// Mitsubishi GX Works2 project: FINAL_V7   PLC: Q03UDV

PROGRAM MAIN
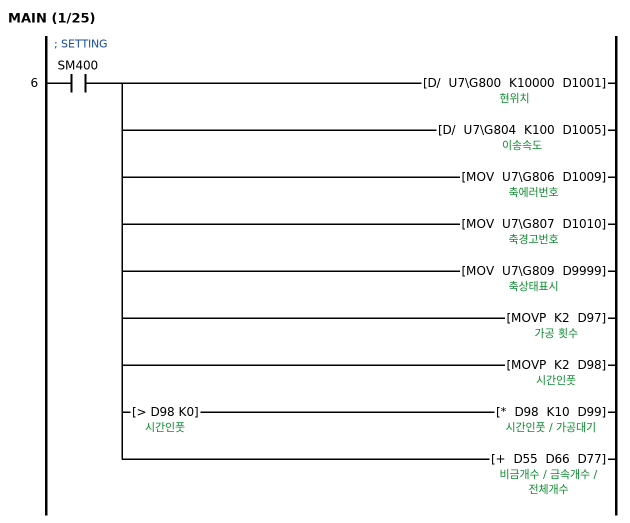
; SETTING
6     LD      SM400
      D/      U7\G800 K10000 D1001  ; 현위치
      D/      U7\G804 K100 D1005  ; 이송속도
      MOV     U7\G806 D1009  ; 축에러번호
      MOV     U7\G807 D1010  ; 축경고번호
      MOV     U7\G809 D9999  ; 축상태표시
      MOVP    K2 D97  ; 가공 횟수
      MOVP    K2 D98  ; 시간인풋
      MPS
      AND>    D98 K0  ; 시간인풋
      *       D98 K10 D99  ; 가공대기
      MPP
      +       D55 D66 D77  ; 비금개수 / 금속개수 / 전체개수
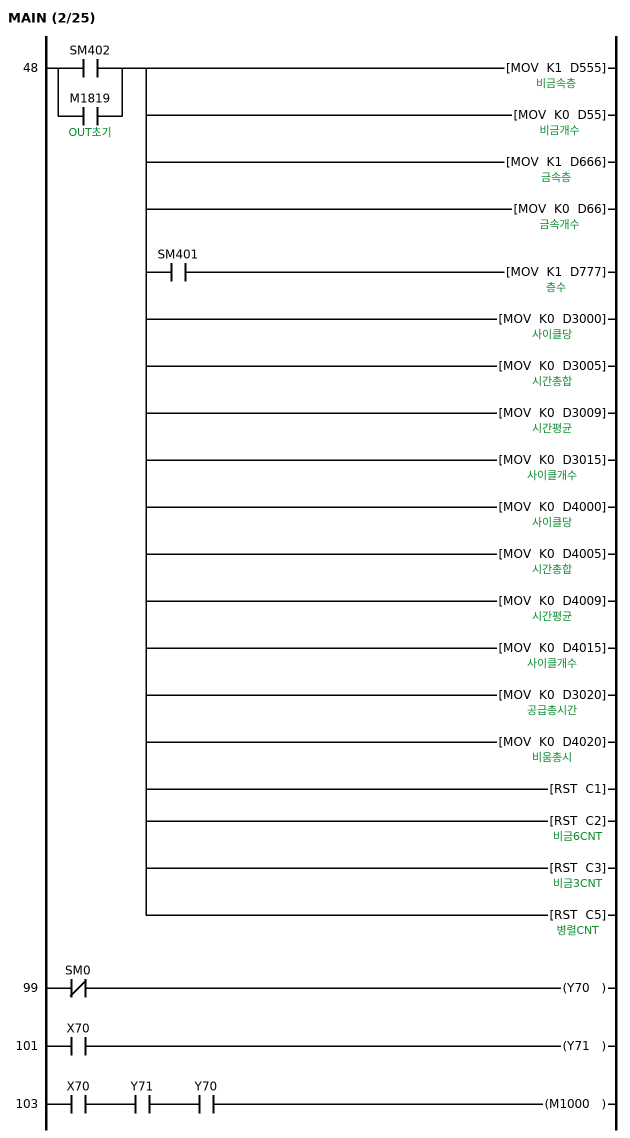
48    LD      SM402
      OR      M1819  ; OUT초기
      MOV     K1 D555  ; 비금속층
      MOV     K0 D55
      MOV     K1 D666  ; 금속층
      MOV     K0 D66
      MPS
      AND     SM401
      MOV     K1 D777  ; 층수
      MPP
      MOV     K0 D3000  ; 사이클당
      MOV     K0 D3005  ; 시간총합
      MOV     K0 D3009  ; 시간평균
      MOV     K0 D3015  ; 사이클개수
      MOV     K0 D4000  ; 사이클당
      MOV     K0 D4005  ; 시간총합
      MOV     K0 D4009  ; 시간평균
      MOV     K0 D4015  ; 사이클개수
      MOV     K0 D3020  ; 공급총시간
      MOV     K0 D4020  ; 비움총시
      RST     C1
      RST     C2  ; 비금6CNT
      RST     C3  ; 비금3CNT
      RST     C5  ; 병렬CNT
99    LDI     SM0
      OUT     Y70
101   LD      X70
      OUT     Y71
103   LD      X70
      AND     Y71
      AND     Y70
      OUT     M1000
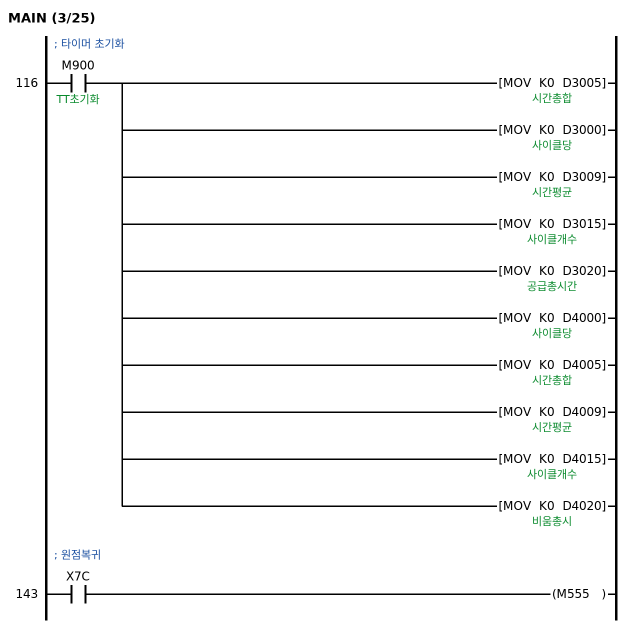
; 타이머 초기화
116   LD      M900  ; TT초기화
      MOV     K0 D3005
      MOV     K0 D3000
      MOV     K0 D3009
      MOV     K0 D3015
      MOV     K0 D3020
      MOV     K0 D4000
      MOV     K0 D4005
      MOV     K0 D4009
      MOV     K0 D4015
      MOV     K0 D4020
; 원점복귀
143   LD      X7C
      OUT     M555
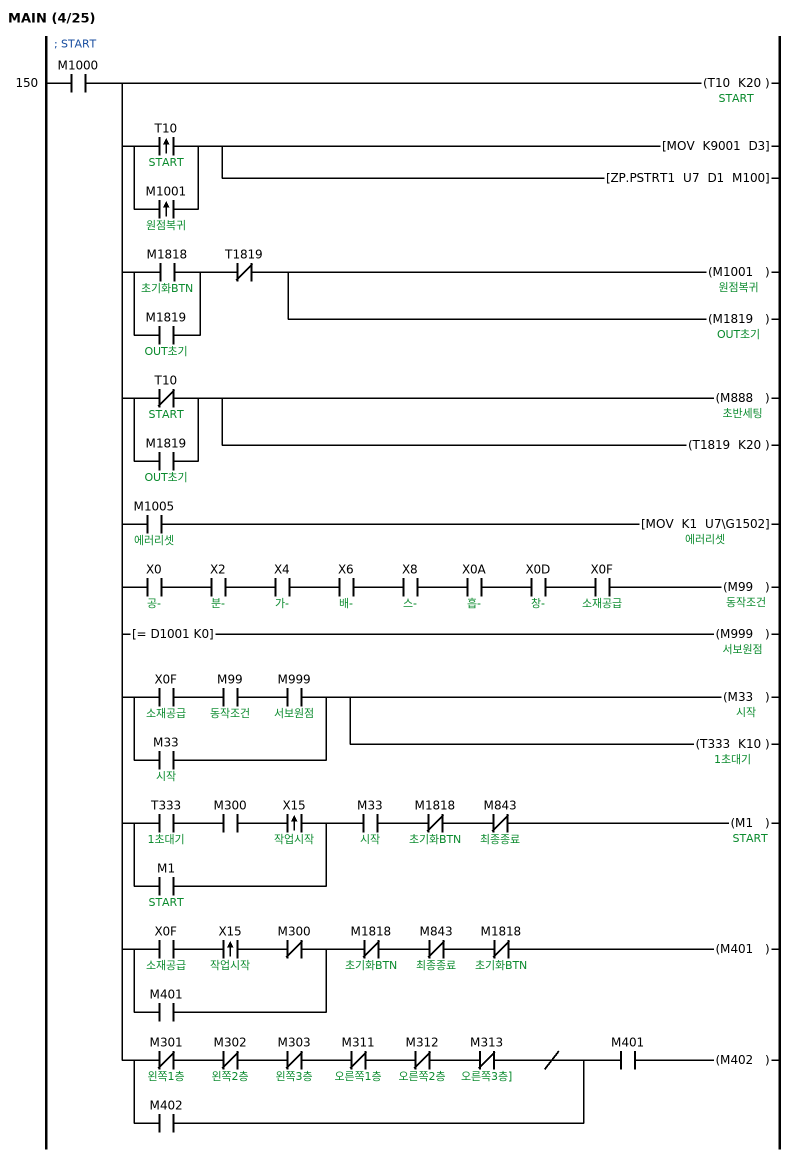
; START
150   LD      M1000
      OUT     T10 K20  ; START
      MPS
      LDP     T10  ; START
      ORP     M1001  ; 원점복귀
      ANB
      MOV     K9001 D3
      ZP.PSTRT1 U7 D1 M100
      MRD
      LD      M1818  ; 초기화BTN
      OR      M1819  ; OUT초기
      ANB
      ANI     T1819
      OUT     M1001  ; 원점복귀
      OUT     M1819  ; OUT초기
      MRD
      LDI     T10  ; START
      OR      M1819  ; OUT초기
      ANB
      OUT     M888  ; 초반세팅
      OUT     T1819 K20
      MRD
      AND     M1005  ; 에러리셋
      MOV     K1 U7\G1502  ; 에러리셋
      MRD
      AND     X0  ; 공-
      AND     X2  ; 분-
      AND     X4  ; 가-
      AND     X6  ; 배-
      AND     X8  ; 스-
      AND     X0A  ; 흡-
      AND     X0D  ; 창-
      AND     X0F  ; 소재공급
      OUT     M99  ; 동작조건
      MRD
      AND=    D1001 K0
      OUT     M999  ; 서보원점
      MRD
      LD      X0F  ; 소재공급
      AND     M99  ; 동작조건
      AND     M999  ; 서보원점
      OR      M33  ; 시작
      ANB
      OUT     M33  ; 시작
      OUT     T333 K10  ; 1초대기
      MRD
      LD      T333  ; 1초대기
      AND     M300
      ANDP    X15  ; 작업시작
      OR      M1  ; START
      ANB
      AND     M33  ; 시작
      ANI     M1818  ; 초기화BTN
      ANI     M843  ; 최종종료
      OUT     M1  ; START
      MRD
      LD      X0F  ; 소재공급
      ANDP    X15  ; 작업시작
      ANI     M300
      OR      M401
      ANB
      ANI     M1818  ; 초기화BTN
      ANI     M843  ; 최종종료
      ANI     M1818  ; 초기화BTN
      OUT     M401
      MPP
      LDI     M301  ; 왼쪽1층
      ANI     M302  ; 왼쪽2층
      ANI     M303  ; 왼쪽3층
      ANI     M311  ; 오른쪽1층
      ANI     M312  ; 오른쪽2층
      ANI     M313  ; 오른쪽3층]
      INV
      OR      M402
      ANB
      AND     M401
      OUT     M402
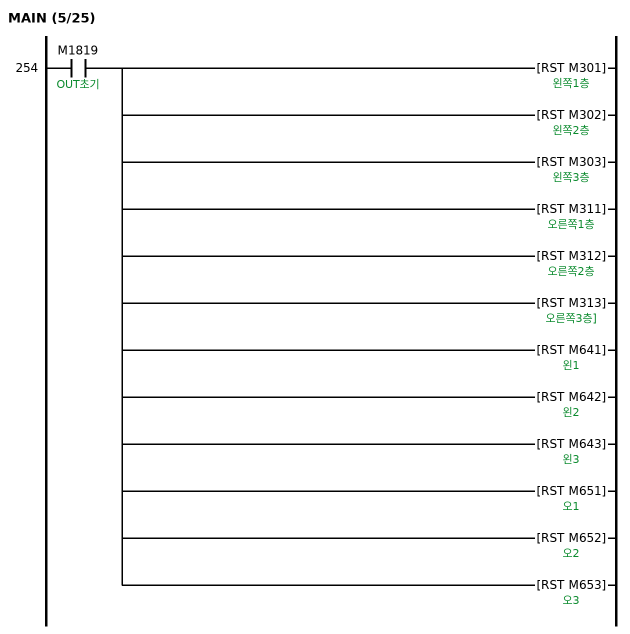
254   LD      M1819  ; OUT초기
      RST     M301  ; 왼쪽1층
      RST     M302  ; 왼쪽2층
      RST     M303  ; 왼쪽3층
      RST     M311  ; 오른쪽1층
      RST     M312  ; 오른쪽2층
      RST     M313  ; 오른쪽3층]
      RST     M641  ; 왼1
      RST     M642  ; 왼2
      RST     M643  ; 왼3
      RST     M651  ; 오1
      RST     M652  ; 오2
      RST     M653  ; 오3
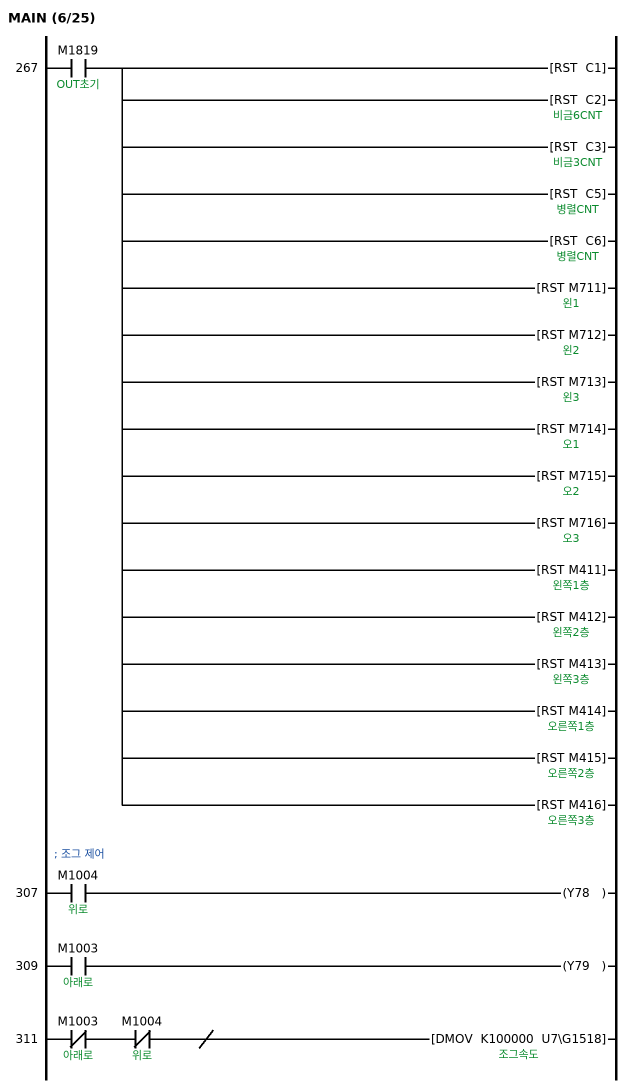
267   LD      M1819  ; OUT초기
      RST     C1
      RST     C2  ; 비금6CNT
      RST     C3  ; 비금3CNT
      RST     C5  ; 병렬CNT
      RST     C6  ; 병렬CNT
      RST     M711  ; 왼1
      RST     M712  ; 왼2
      RST     M713  ; 왼3
      RST     M714  ; 오1
      RST     M715  ; 오2
      RST     M716  ; 오3
      RST     M411  ; 왼쪽1층
      RST     M412  ; 왼쪽2층
      RST     M413  ; 왼쪽3층
      RST     M414  ; 오른쪽1층
      RST     M415  ; 오른쪽2층
      RST     M416  ; 오른쪽3층
; 조그 제어
307   LD      M1004  ; 위로
      OUT     Y78
309   LD      M1003  ; 아래로
      OUT     Y79
311   LDI     M1003  ; 아래로
      ANI     M1004  ; 위로
      INV
      DMOV    K100000 U7\G1518  ; 조그속도
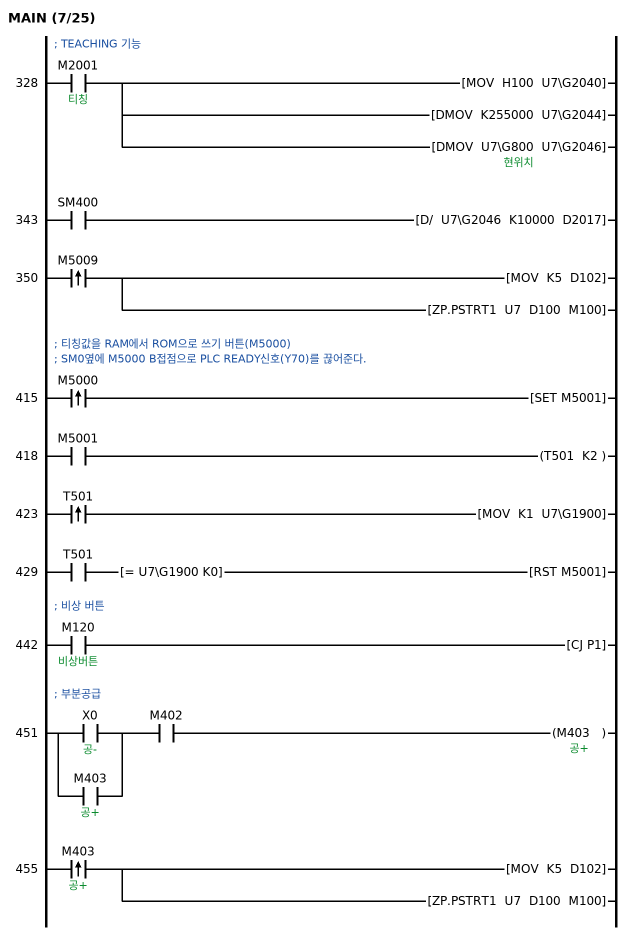
; TEACHING 기능
328   LD      M2001  ; 티칭
      MOV     H100 U7\G2040
      DMOV    K255000 U7\G2044
      DMOV    U7\G800 U7\G2046
343   LD      SM400
      D/      U7\G2046 K10000 D2017
350   LDP     M5009
      MOV     K5 D102
      ZP.PSTRT1 U7 D100 M100
; 티칭값을 RAM에서 ROM으로 쓰기 버튼(M5000)
; SM0옆에 M5000 B접점으로 PLC READY신호(Y70)를 끊어준다.
415   LDP     M5000
      SET     M5001
418   LD      M5001
      OUT     T501 K2
423   LDP     T501
      MOV     K1 U7\G1900
429   LD      T501
      AND=    U7\G1900 K0
      RST     M5001
; 비상 버튼
442   LD      M120  ; 비상버튼
      CJ      P1
; 부분공급
451   LD      X0  ; 공-
      OR      M403  ; 공+
      AND     M402
      OUT     M403  ; 공+
455   LDP     M403  ; 공+
      MOV     K5 D102
      ZP.PSTRT1 U7 D100 M100
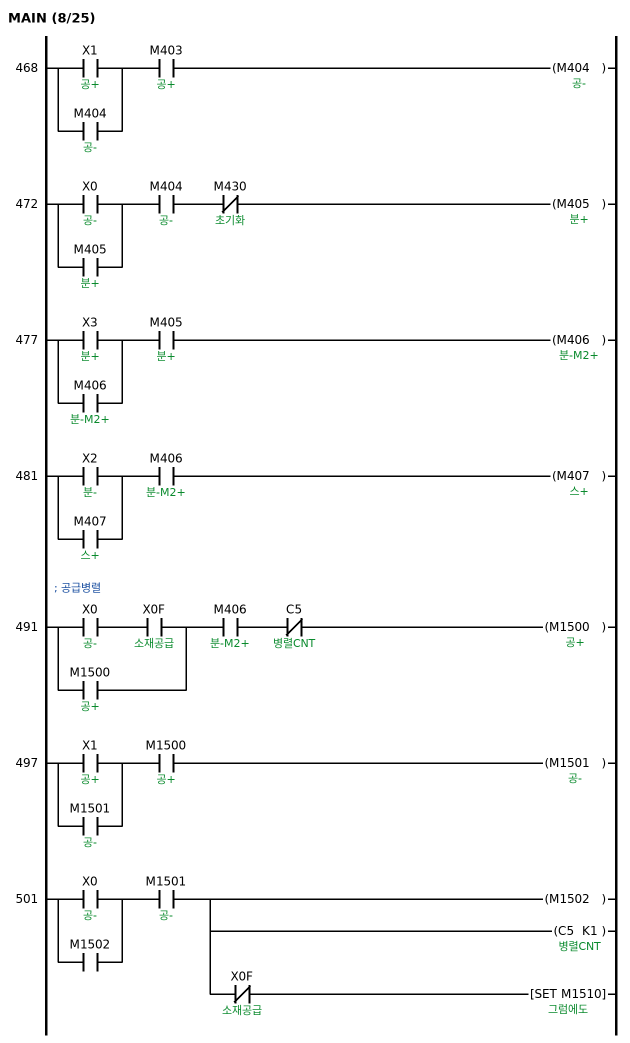
468   LD      X1  ; 공+
      OR      M404  ; 공-
      AND     M403  ; 공+
      OUT     M404  ; 공-
472   LD      X0  ; 공-
      OR      M405  ; 분+
      AND     M404  ; 공-
      ANI     M430  ; 초기화
      OUT     M405  ; 분+
477   LD      X3  ; 분+
      OR      M406  ; 분-M2+
      AND     M405  ; 분+
      OUT     M406  ; 분-M2+
481   LD      X2  ; 분-
      OR      M407  ; 스+
      AND     M406  ; 분-M2+
      OUT     M407  ; 스+
; 공급병렬
491   LD      X0  ; 공-
      AND     X0F  ; 소재공급
      OR      M1500  ; 공+
      AND     M406  ; 분-M2+
      ANI     C5  ; 병렬CNT
      OUT     M1500  ; 공+
497   LD      X1  ; 공+
      OR      M1501  ; 공-
      AND     M1500  ; 공+
      OUT     M1501  ; 공-
501   LD      X0  ; 공-
      OR      M1502
      AND     M1501  ; 공-
      OUT     M1502
      OUT     C5 K1  ; 병렬CNT
      ANI     X0F  ; 소재공급
      SET     M1510  ; 그럼에도
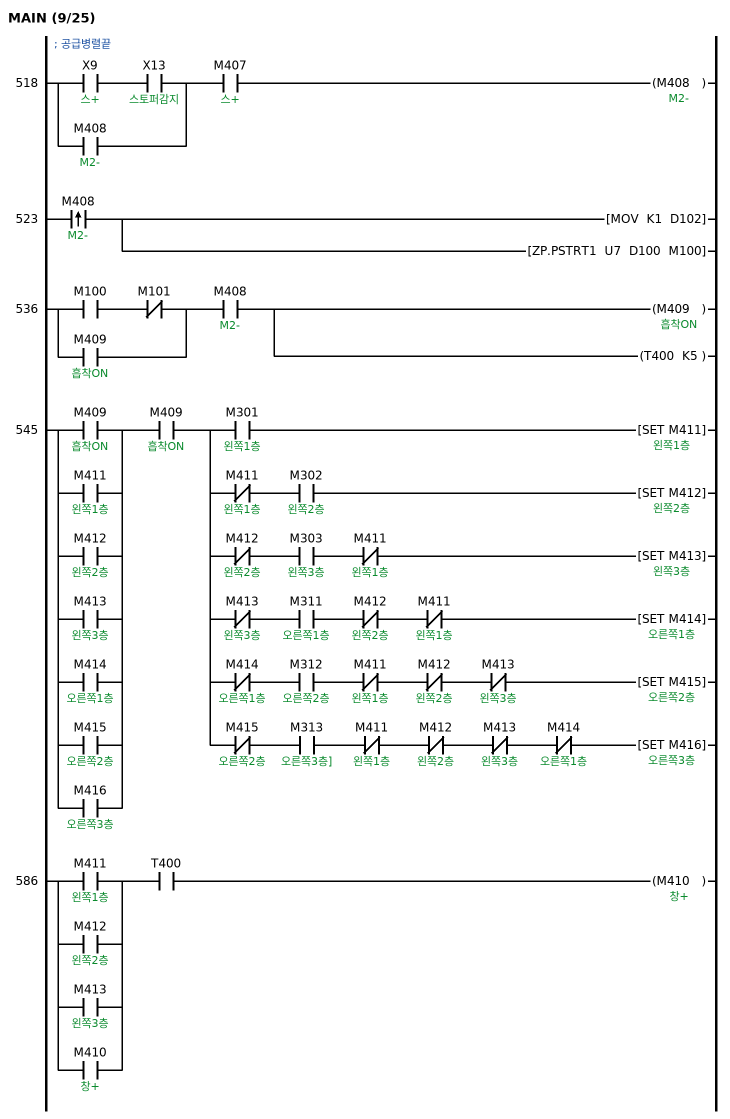
; 공급병렬끝
518   LD      X9  ; 스+
      AND     X13  ; 스토퍼감지
      OR      M408  ; M2-
      AND     M407  ; 스+
      OUT     M408  ; M2-
523   LDP     M408  ; M2-
      MOV     K1 D102
      ZP.PSTRT1 U7 D100 M100
536   LD      M100
      ANI     M101
      OR      M409  ; 흡착ON
      AND     M408  ; M2-
      OUT     M409  ; 흡착ON
      OUT     T400 K5
545   LD      M409  ; 흡착ON
      OR      M411  ; 왼쪽1층
      OR      M412  ; 왼쪽2층
      OR      M413  ; 왼쪽3층
      OR      M414  ; 오른쪽1층
      OR      M415  ; 오른쪽2층
      OR      M416  ; 오른쪽3층
      AND     M409  ; 흡착ON
      MPS
      AND     M301  ; 왼쪽1층
      SET     M411  ; 왼쪽1층
      MRD
      ANI     M411  ; 왼쪽1층
      AND     M302  ; 왼쪽2층
      SET     M412  ; 왼쪽2층
      MRD
      ANI     M412  ; 왼쪽2층
      AND     M303  ; 왼쪽3층
      ANI     M411  ; 왼쪽1층
      SET     M413  ; 왼쪽3층
      MRD
      ANI     M413  ; 왼쪽3층
      AND     M311  ; 오른쪽1층
      ANI     M412  ; 왼쪽2층
      ANI     M411  ; 왼쪽1층
      SET     M414  ; 오른쪽1층
      MRD
      ANI     M414  ; 오른쪽1층
      AND     M312  ; 오른쪽2층
      ANI     M411  ; 왼쪽1층
      ANI     M412  ; 왼쪽2층
      ANI     M413  ; 왼쪽3층
      SET     M415  ; 오른쪽2층
      MPP
      ANI     M415  ; 오른쪽2층
      AND     M313  ; 오른쪽3층]
      ANI     M411  ; 왼쪽1층
      ANI     M412  ; 왼쪽2층
      ANI     M413  ; 왼쪽3층
      ANI     M414  ; 오른쪽1층
      SET     M416  ; 오른쪽3층
586   LD      M411  ; 왼쪽1층
      OR      M412  ; 왼쪽2층
      OR      M413  ; 왼쪽3층
      OR      M410  ; 창+
      AND     T400
      OUT     M410  ; 창+
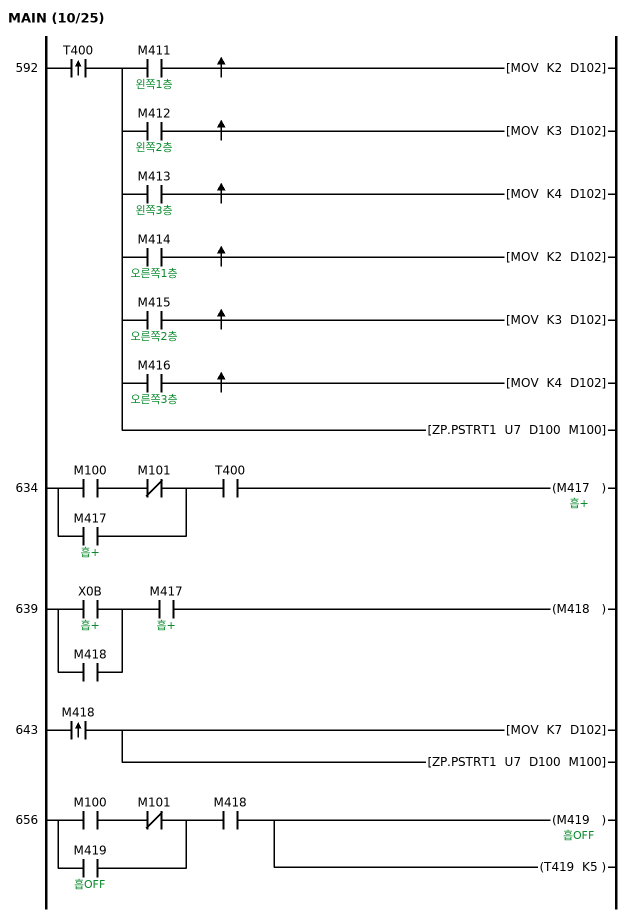
592   LDP     T400
      MPS
      AND     M411  ; 왼쪽1층
      MEP
      MOV     K2 D102
      MRD
      AND     M412  ; 왼쪽2층
      MEP
      MOV     K3 D102
      MRD
      AND     M413  ; 왼쪽3층
      MEP
      MOV     K4 D102
      MRD
      AND     M414  ; 오른쪽1층
      MEP
      MOV     K2 D102
      MRD
      AND     M415  ; 오른쪽2층
      MEP
      MOV     K3 D102
      MRD
      AND     M416  ; 오른쪽3층
      MEP
      MOV     K4 D102
      MPP
      ZP.PSTRT1 U7 D100 M100
634   LD      M100
      ANI     M101
      OR      M417  ; 흡+
      AND     T400
      OUT     M417  ; 흡+
639   LD      X0B  ; 흡+
      OR      M418
      AND     M417  ; 흡+
      OUT     M418
643   LDP     M418
      MOV     K7 D102
      ZP.PSTRT1 U7 D100 M100
656   LD      M100
      ANI     M101
      OR      M419  ; 흡OFF
      AND     M418
      OUT     M419  ; 흡OFF
      OUT     T419 K5
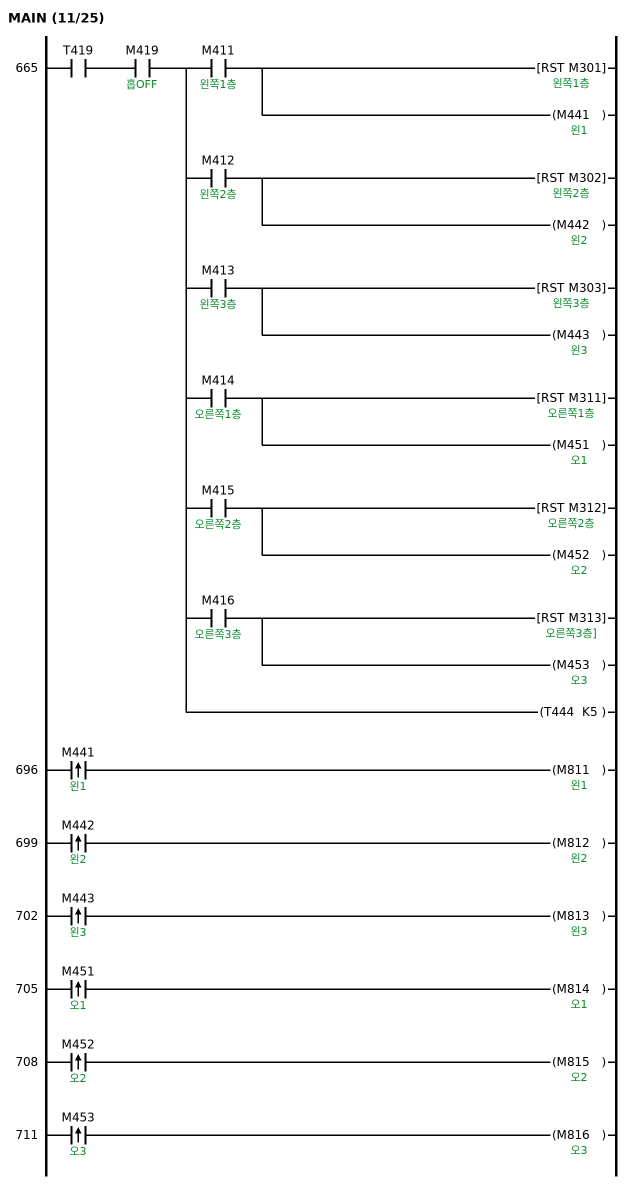
665   LD      T419
      AND     M419  ; 흡OFF
      MPS
      AND     M411  ; 왼쪽1층
      RST     M301  ; 왼쪽1층
      OUT     M441  ; 왼1
      MRD
      AND     M412  ; 왼쪽2층
      RST     M302  ; 왼쪽2층
      OUT     M442  ; 왼2
      MRD
      AND     M413  ; 왼쪽3층
      RST     M303  ; 왼쪽3층
      OUT     M443  ; 왼3
      MRD
      AND     M414  ; 오른쪽1층
      RST     M311  ; 오른쪽1층
      OUT     M451  ; 오1
      MRD
      AND     M415  ; 오른쪽2층
      RST     M312  ; 오른쪽2층
      OUT     M452  ; 오2
      MRD
      AND     M416  ; 오른쪽3층
      RST     M313  ; 오른쪽3층]
      OUT     M453  ; 오3
      MPP
      OUT     T444 K5
696   LDP     M441  ; 왼1
      OUT     M811  ; 왼1
699   LDP     M442  ; 왼2
      OUT     M812  ; 왼2
702   LDP     M443  ; 왼3
      OUT     M813  ; 왼3
705   LDP     M451  ; 오1
      OUT     M814  ; 오1
708   LDP     M452  ; 오2
      OUT     M815  ; 오2
711   LDP     M453  ; 오3
      OUT     M816  ; 오3
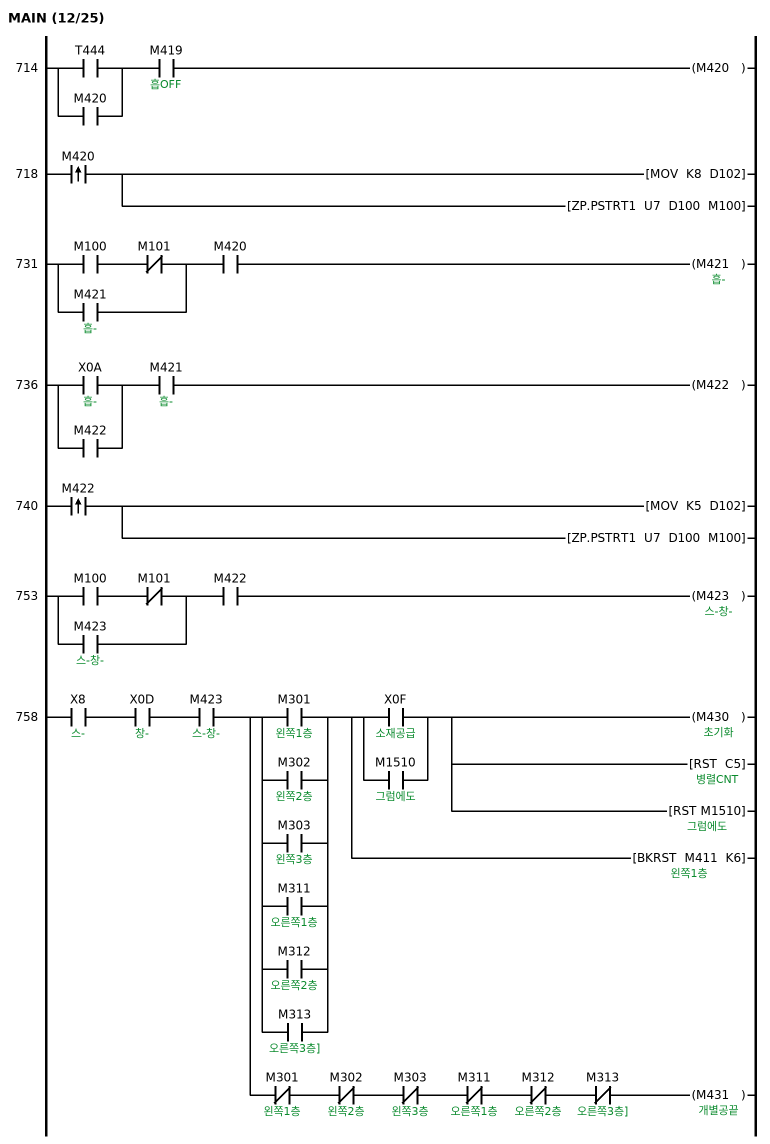
714   LD      T444
      OR      M420
      AND     M419  ; 흡OFF
      OUT     M420
718   LDP     M420
      MOV     K8 D102
      ZP.PSTRT1 U7 D100 M100
731   LD      M100
      ANI     M101
      OR      M421  ; 흡-
      AND     M420
      OUT     M421  ; 흡-
736   LD      X0A  ; 흡-
      OR      M422
      AND     M421  ; 흡-
      OUT     M422
740   LDP     M422
      MOV     K5 D102
      ZP.PSTRT1 U7 D100 M100
753   LD      M100
      ANI     M101
      OR      M423  ; 스-창-
      AND     M422
      OUT     M423  ; 스-창-
758   LD      X8  ; 스-
      AND     X0D  ; 창-
      AND     M423  ; 스-창-
      MPS
      LD      M301  ; 왼쪽1층
      OR      M302  ; 왼쪽2층
      OR      M303  ; 왼쪽3층
      OR      M311  ; 오른쪽1층
      OR      M312  ; 오른쪽2층
      OR      M313  ; 오른쪽3층]
      ANB
      MPS
      LD      X0F  ; 소재공급
      OR      M1510  ; 그럼에도
      ANB
      OUT     M430  ; 초기화
      RST     C5  ; 병렬CNT
      RST     M1510  ; 그럼에도
      MPP
      BKRST   M411 K6
      MPP
      ANI     M301  ; 왼쪽1층
      ANI     M302  ; 왼쪽2층
      ANI     M303  ; 왼쪽3층
      ANI     M311  ; 오른쪽1층
      ANI     M312  ; 오른쪽2층
      ANI     M313  ; 오른쪽3층]
      OUT     M431  ; 개별공끝
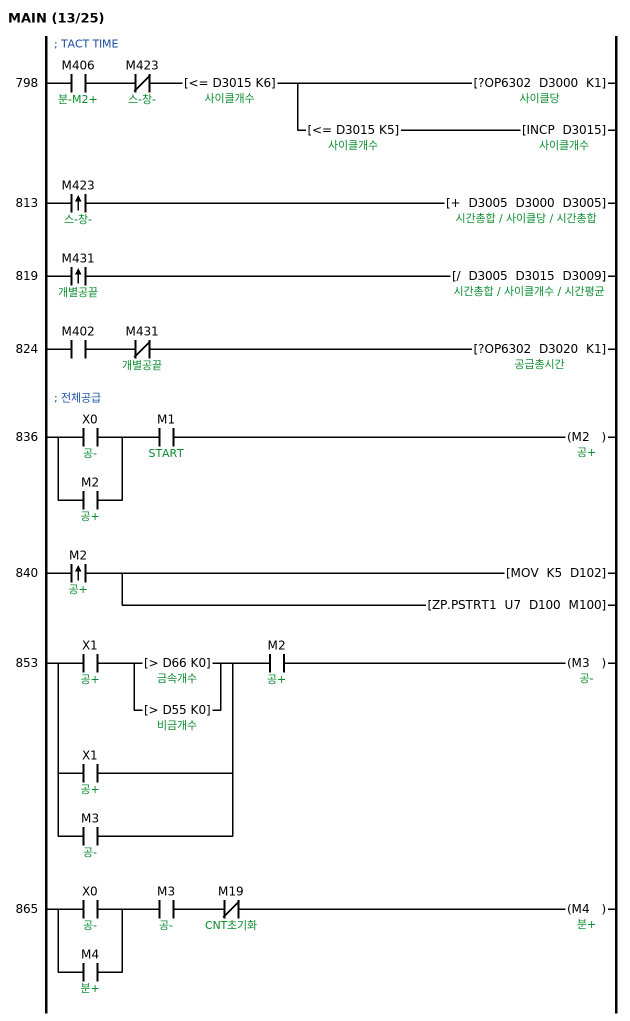
; TACT TIME
798   LD      M406  ; 분-M2+
      ANI     M423  ; 스-창-
      AND<=   D3015 K6  ; 사이클개수
      ?OP6302 D3000 K1
      AND<=   D3015 K5  ; 사이클개수
      INCP    D3015
813   LDP     M423  ; 스-창-
      +       D3005 D3000 D3005
819   LDP     M431  ; 개별공끝
      /       D3005 D3015 D3009
824   LD      M402
      ANI     M431  ; 개별공끝
      ?OP6302 D3020 K1
; 전체공급
836   LD      X0  ; 공-
      OR      M2  ; 공+
      AND     M1  ; START
      OUT     M2  ; 공+
840   LDP     M2  ; 공+
      MOV     K5 D102
      ZP.PSTRT1 U7 D100 M100
853   LD      X1  ; 공+
      LD>     D66 K0  ; 금속개수
      OR>     D55 K0  ; 비금개수
      ANB
      OR      X1  ; 공+
      OR      M3  ; 공-
      AND     M2  ; 공+
      OUT     M3  ; 공-
865   LD      X0  ; 공-
      OR      M4  ; 분+
      AND     M3  ; 공-
      ANI     M19  ; CNT초기화
      OUT     M4  ; 분+
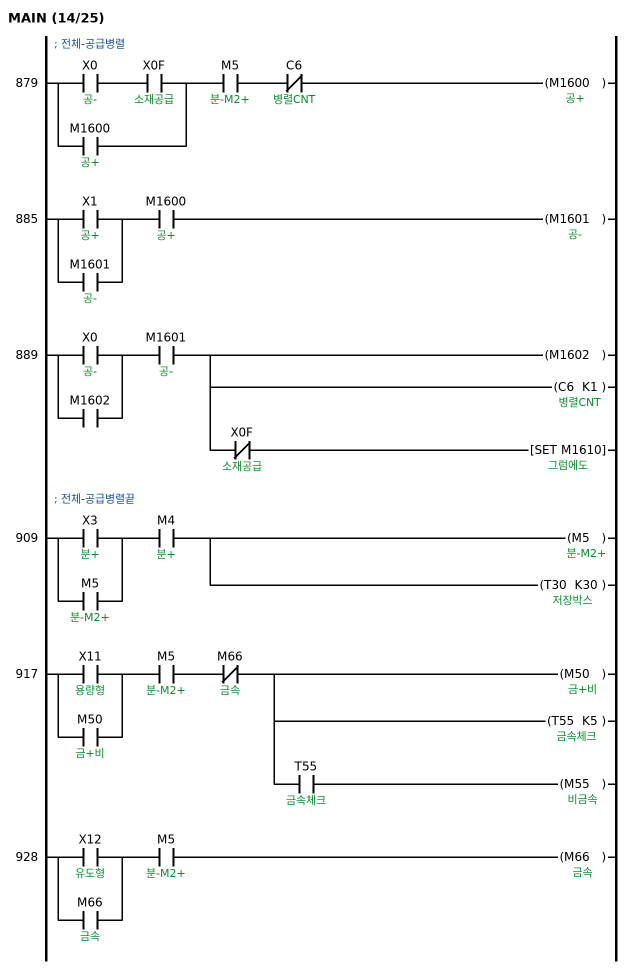
; 전체-공급병렬
879   LD      X0  ; 공-
      AND     X0F  ; 소재공급
      OR      M1600  ; 공+
      AND     M5  ; 분-M2+
      ANI     C6  ; 병렬CNT
      OUT     M1600  ; 공+
885   LD      X1  ; 공+
      OR      M1601  ; 공-
      AND     M1600  ; 공+
      OUT     M1601  ; 공-
889   LD      X0  ; 공-
      OR      M1602
      AND     M1601  ; 공-
      OUT     M1602
      OUT     C6 K1  ; 병렬CNT
      ANI     X0F  ; 소재공급
      SET     M1610  ; 그럼에도
; 전체-공급병렬끝
909   LD      X3  ; 분+
      OR      M5  ; 분-M2+
      AND     M4  ; 분+
      OUT     M5  ; 분-M2+
      OUT     T30 K30  ; 저장박스
917   LD      X11  ; 용량형
      OR      M50  ; 금+비
      AND     M5  ; 분-M2+
      ANI     M66  ; 금속
      OUT     M50  ; 금+비
      OUT     T55 K5  ; 금속체크
      AND     T55  ; 금속체크
      OUT     M55  ; 비금속
928   LD      X12  ; 유도형
      OR      M66  ; 금속
      AND     M5  ; 분-M2+
      OUT     M66  ; 금속
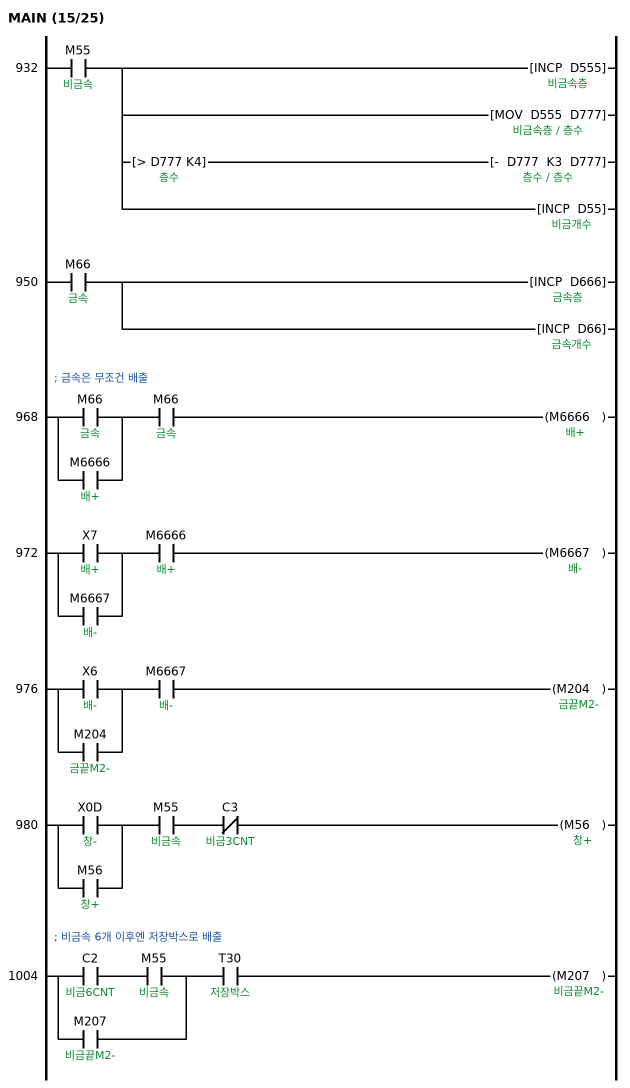
932   LD      M55  ; 비금속
      INCP    D555
      MOV     D555 D777
      MPS
      AND>    D777 K4  ; 층수
      -       D777 K3 D777
      MPP
      INCP    D55
950   LD      M66  ; 금속
      INCP    D666
      INCP    D66
; 금속은 무조건 배출
968   LD      M66  ; 금속
      OR      M6666  ; 배+
      AND     M66  ; 금속
      OUT     M6666  ; 배+
972   LD      X7  ; 배+
      OR      M6667  ; 배-
      AND     M6666  ; 배+
      OUT     M6667  ; 배-
976   LD      X6  ; 배-
      OR      M204  ; 금끝M2-
      AND     M6667  ; 배-
      OUT     M204  ; 금끝M2-
980   LD      X0D  ; 창-
      OR      M56  ; 창+
      AND     M55  ; 비금속
      ANI     C3  ; 비금3CNT
      OUT     M56  ; 창+
; 비금속 6개 이후엔 저장박스로 배출
1004  LD      C2  ; 비금6CNT
      AND     M55  ; 비금속
      OR      M207  ; 비금끝M2-
      AND     T30  ; 저장박스
      OUT     M207  ; 비금끝M2-
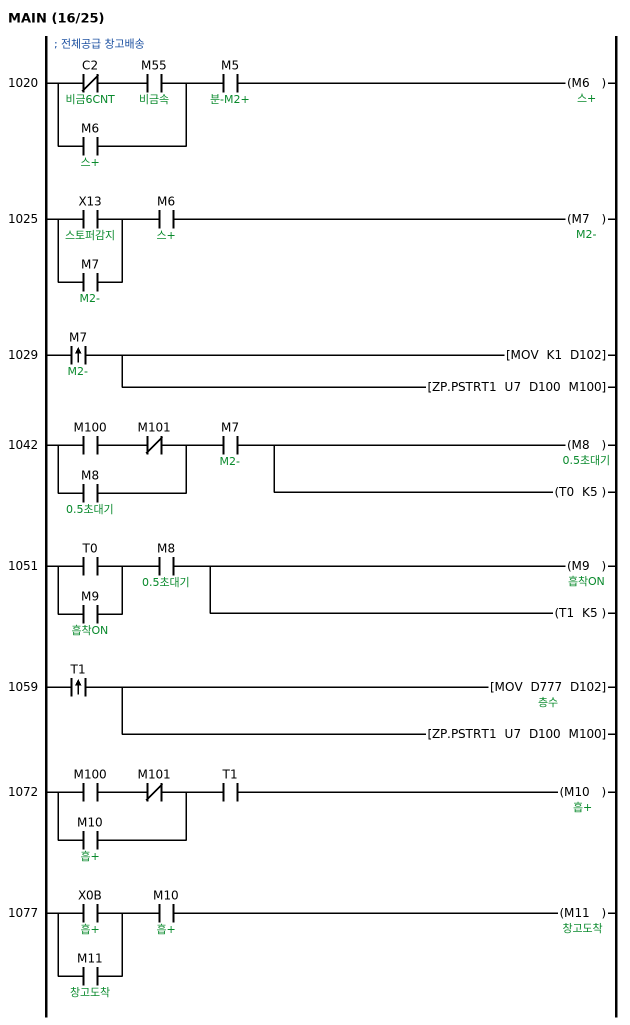
; 전체공급 창고배송
1020  LDI     C2  ; 비금6CNT
      AND     M55  ; 비금속
      OR      M6  ; 스+
      AND     M5  ; 분-M2+
      OUT     M6  ; 스+
1025  LD      X13  ; 스토퍼감지
      OR      M7  ; M2-
      AND     M6  ; 스+
      OUT     M7  ; M2-
1029  LDP     M7  ; M2-
      MOV     K1 D102
      ZP.PSTRT1 U7 D100 M100
1042  LD      M100
      ANI     M101
      OR      M8  ; 0.5초대기
      AND     M7  ; M2-
      OUT     M8  ; 0.5초대기
      OUT     T0 K5
1051  LD      T0
      OR      M9  ; 흡착ON
      AND     M8  ; 0.5초대기
      OUT     M9  ; 흡착ON
      OUT     T1 K5
1059  LDP     T1
      MOV     D777 D102
      ZP.PSTRT1 U7 D100 M100
1072  LD      M100
      ANI     M101
      OR      M10  ; 흡+
      AND     T1
      OUT     M10  ; 흡+
1077  LD      X0B  ; 흡+
      OR      M11  ; 창고도착
      AND     M10  ; 흡+
      OUT     M11  ; 창고도착
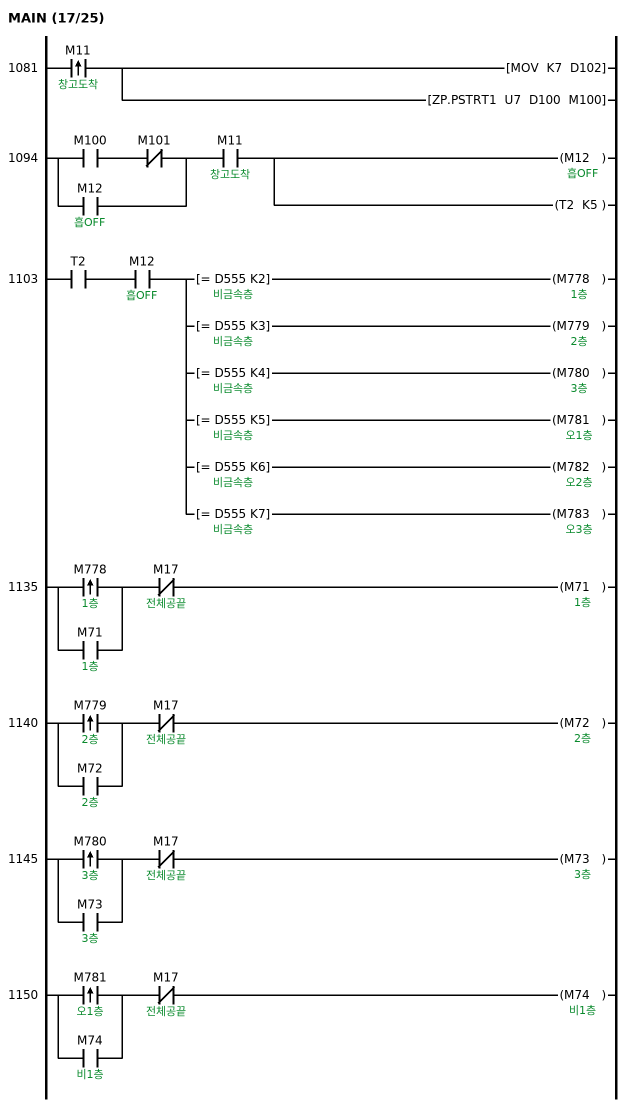
1081  LDP     M11  ; 창고도착
      MOV     K7 D102
      ZP.PSTRT1 U7 D100 M100
1094  LD      M100
      ANI     M101
      OR      M12  ; 흡OFF
      AND     M11  ; 창고도착
      OUT     M12  ; 흡OFF
      OUT     T2 K5
1103  LD      T2
      AND     M12  ; 흡OFF
      MPS
      AND=    D555 K2  ; 비금속층
      OUT     M778  ; 1층
      MRD
      AND=    D555 K3  ; 비금속층
      OUT     M779  ; 2층
      MRD
      AND=    D555 K4  ; 비금속층
      OUT     M780  ; 3층
      MRD
      AND=    D555 K5  ; 비금속층
      OUT     M781  ; 오1층
      MRD
      AND=    D555 K6  ; 비금속층
      OUT     M782  ; 오2층
      MPP
      AND=    D555 K7  ; 비금속층
      OUT     M783  ; 오3층
1135  LDP     M778  ; 1층
      OR      M71  ; 1층
      ANI     M17  ; 전체공끝
      OUT     M71  ; 1층
1140  LDP     M779  ; 2층
      OR      M72  ; 2층
      ANI     M17  ; 전체공끝
      OUT     M72  ; 2층
1145  LDP     M780  ; 3층
      OR      M73  ; 3층
      ANI     M17  ; 전체공끝
      OUT     M73  ; 3층
1150  LDP     M781  ; 오1층
      OR      M74  ; 비1층
      ANI     M17  ; 전체공끝
      OUT     M74  ; 비1층
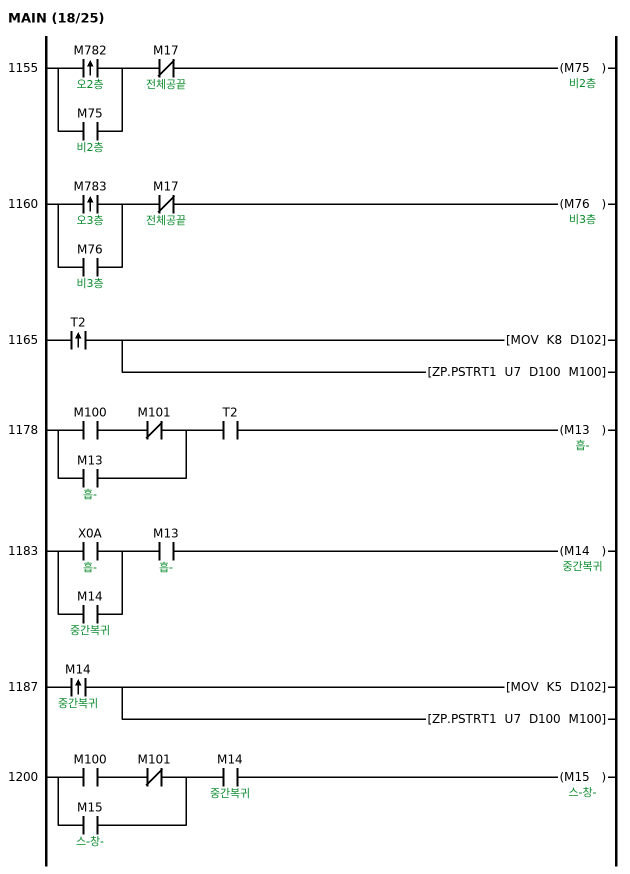
1155  LDP     M782  ; 오2층
      OR      M75  ; 비2층
      ANI     M17  ; 전체공끝
      OUT     M75  ; 비2층
1160  LDP     M783  ; 오3층
      OR      M76  ; 비3층
      ANI     M17  ; 전체공끝
      OUT     M76  ; 비3층
1165  LDP     T2
      MOV     K8 D102
      ZP.PSTRT1 U7 D100 M100
1178  LD      M100
      ANI     M101
      OR      M13  ; 흡-
      AND     T2
      OUT     M13  ; 흡-
1183  LD      X0A  ; 흡-
      OR      M14  ; 중간복귀
      AND     M13  ; 흡-
      OUT     M14  ; 중간복귀
1187  LDP     M14  ; 중간복귀
      MOV     K5 D102
      ZP.PSTRT1 U7 D100 M100
1200  LD      M100
      ANI     M101
      OR      M15  ; 스-창-
      AND     M14  ; 중간복귀
      OUT     M15  ; 스-창-
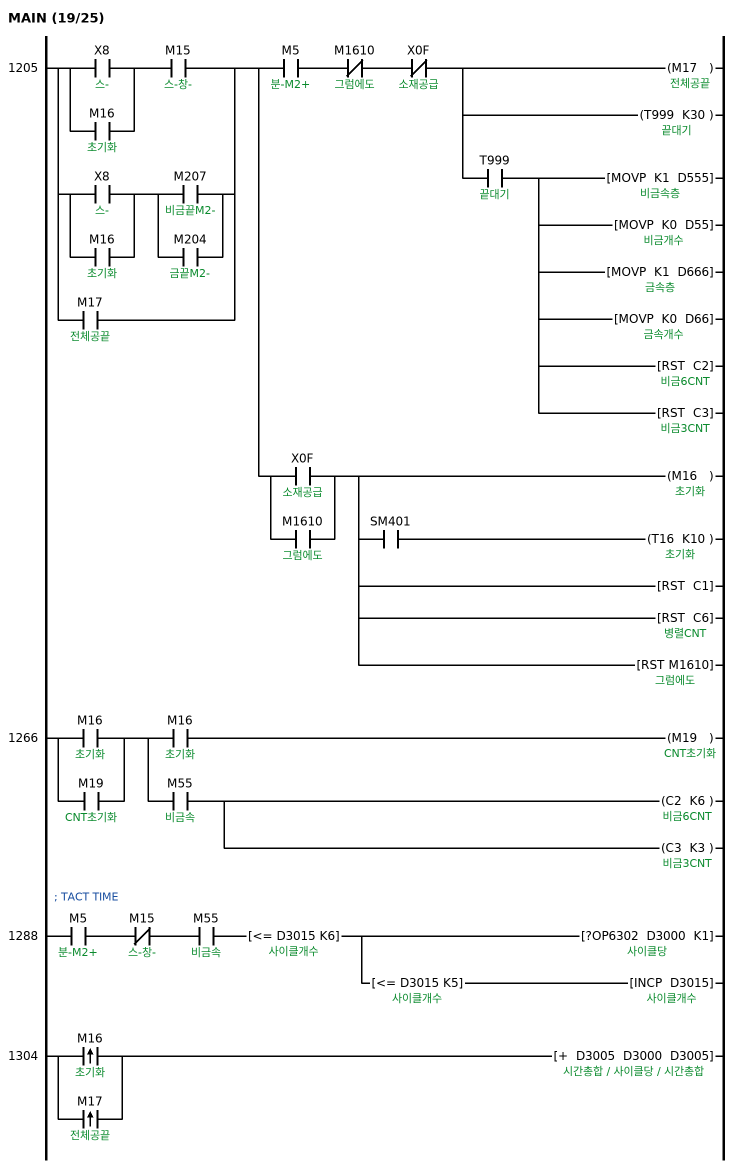
1205  LD      X8  ; 스-
      OR      M16  ; 초기화
      AND     M15  ; 스-창-
      LD      X8  ; 스-
      OR      M16  ; 초기화
      LD      M207  ; 비금끝M2-
      OR      M204  ; 금끝M2-
      ANB
      ORB
      OR      M17  ; 전체공끝
      MPS
      AND     M5  ; 분-M2+
      ANI     M1610  ; 그럼에도
      ANI     X0F  ; 소재공급
      OUT     M17  ; 전체공끝
      OUT     T999 K30  ; 끝대기
      AND     T999  ; 끝대기
      MOVP    K1 D555
      MOVP    K0 D55
      MOVP    K1 D666
      MOVP    K0 D66
      RST     C2  ; 비금6CNT
      RST     C3  ; 비금3CNT
      MPP
      LD      X0F  ; 소재공급
      OR      M1610  ; 그럼에도
      ANB
      OUT     M16  ; 초기화
      MPS
      AND     SM401
      OUT     T16 K10  ; 초기화
      MPP
      RST     C1
      RST     C6  ; 병렬CNT
      RST     M1610  ; 그럼에도
1266  LD      M16  ; 초기화
      OR      M19  ; CNT초기화
      MPS
      AND     M16  ; 초기화
      OUT     M19  ; CNT초기화
      MPP
      AND     M55  ; 비금속
      OUT     C2 K6  ; 비금6CNT
      OUT     C3 K3  ; 비금3CNT
; TACT TIME
1288  LD      M5  ; 분-M2+
      ANI     M15  ; 스-창-
      AND     M55  ; 비금속
      AND<=   D3015 K6  ; 사이클개수
      ?OP6302 D3000 K1
      AND<=   D3015 K5  ; 사이클개수
      INCP    D3015
1304  LDP     M16  ; 초기화
      ORP     M17  ; 전체공끝
      +       D3005 D3000 D3005
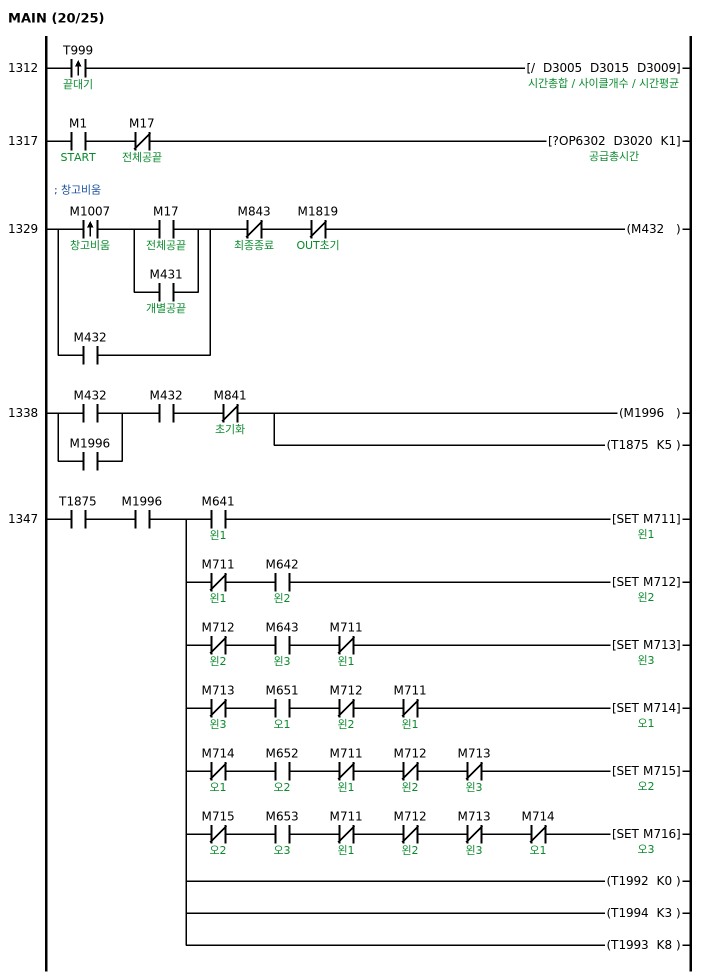
1312  LDP     T999  ; 끝대기
      /       D3005 D3015 D3009
1317  LD      M1  ; START
      ANI     M17  ; 전체공끝
      ?OP6302 D3020 K1
; 창고비움
1329  LDP     M1007  ; 창고비움
      LD      M17  ; 전체공끝
      OR      M431  ; 개별공끝
      ANB
      OR      M432
      ANI     M843  ; 최종종료
      ANI     M1819  ; OUT초기
      OUT     M432
1338  LD      M432
      OR      M1996
      AND     M432
      ANI     M841  ; 초기화
      OUT     M1996
      OUT     T1875 K5
1347  LD      T1875
      AND     M1996
      MPS
      AND     M641  ; 왼1
      SET     M711  ; 왼1
      MRD
      ANI     M711  ; 왼1
      AND     M642  ; 왼2
      SET     M712  ; 왼2
      MRD
      ANI     M712  ; 왼2
      AND     M643  ; 왼3
      ANI     M711  ; 왼1
      SET     M713  ; 왼3
      MRD
      ANI     M713  ; 왼3
      AND     M651  ; 오1
      ANI     M712  ; 왼2
      ANI     M711  ; 왼1
      SET     M714  ; 오1
      MRD
      ANI     M714  ; 오1
      AND     M652  ; 오2
      ANI     M711  ; 왼1
      ANI     M712  ; 왼2
      ANI     M713  ; 왼3
      SET     M715  ; 오2
      MRD
      ANI     M715  ; 오2
      AND     M653  ; 오3
      ANI     M711  ; 왼1
      ANI     M712  ; 왼2
      ANI     M713  ; 왼3
      ANI     M714  ; 오1
      SET     M716  ; 오3
      MPP
      OUT     T1992 K0
      OUT     T1994 K3
      OUT     T1993 K8
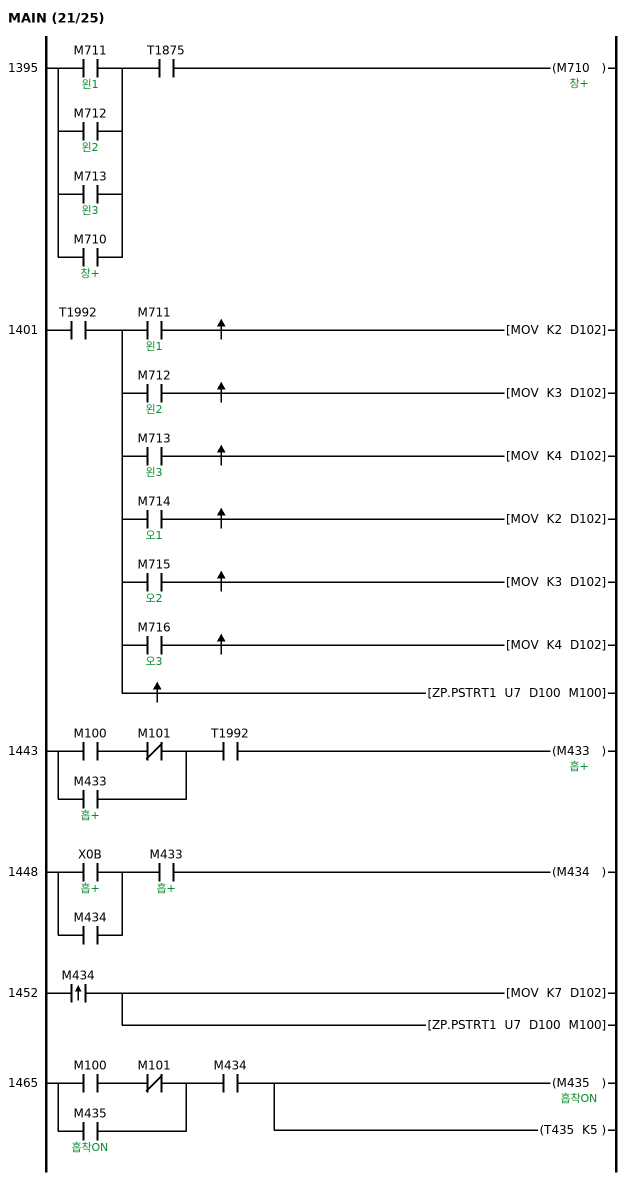
1395  LD      M711  ; 왼1
      OR      M712  ; 왼2
      OR      M713  ; 왼3
      OR      M710  ; 창+
      AND     T1875
      OUT     M710  ; 창+
1401  LD      T1992
      MPS
      AND     M711  ; 왼1
      MEP
      MOV     K2 D102
      MRD
      AND     M712  ; 왼2
      MEP
      MOV     K3 D102
      MRD
      AND     M713  ; 왼3
      MEP
      MOV     K4 D102
      MRD
      AND     M714  ; 오1
      MEP
      MOV     K2 D102
      MRD
      AND     M715  ; 오2
      MEP
      MOV     K3 D102
      MRD
      AND     M716  ; 오3
      MEP
      MOV     K4 D102
      MPP
      MEP
      ZP.PSTRT1 U7 D100 M100
1443  LD      M100
      ANI     M101
      OR      M433  ; 흡+
      AND     T1992
      OUT     M433  ; 흡+
1448  LD      X0B  ; 흡+
      OR      M434
      AND     M433  ; 흡+
      OUT     M434
1452  LDP     M434
      MOV     K7 D102
      ZP.PSTRT1 U7 D100 M100
1465  LD      M100
      ANI     M101
      OR      M435  ; 흡착ON
      AND     M434
      OUT     M435  ; 흡착ON
      OUT     T435 K5
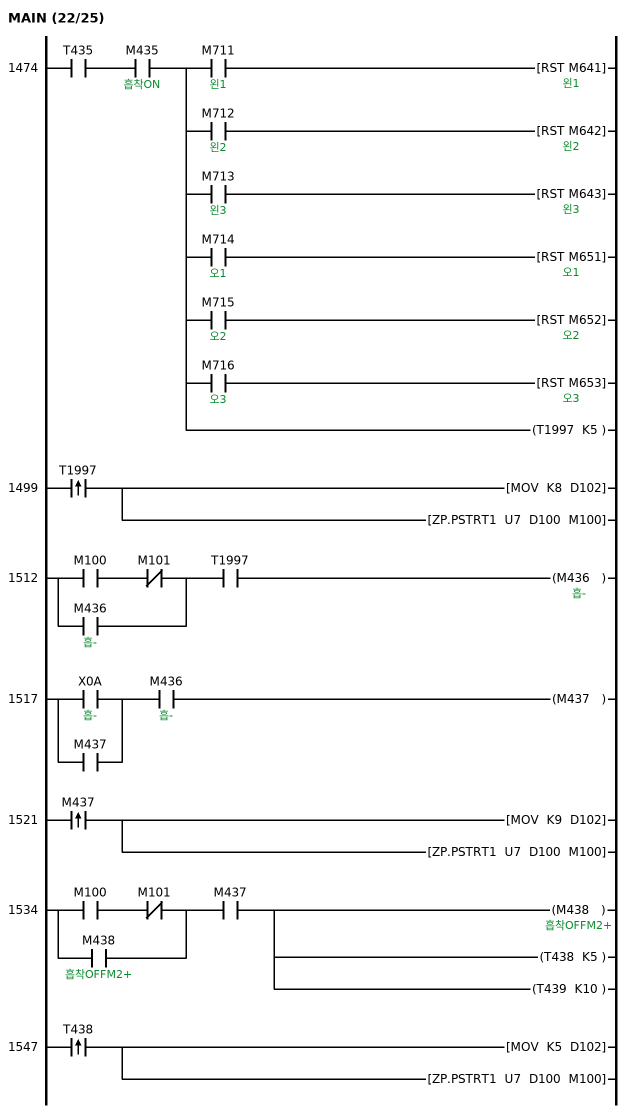
1474  LD      T435
      AND     M435  ; 흡착ON
      MPS
      AND     M711  ; 왼1
      RST     M641  ; 왼1
      MRD
      AND     M712  ; 왼2
      RST     M642  ; 왼2
      MRD
      AND     M713  ; 왼3
      RST     M643  ; 왼3
      MRD
      AND     M714  ; 오1
      RST     M651  ; 오1
      MRD
      AND     M715  ; 오2
      RST     M652  ; 오2
      MRD
      AND     M716  ; 오3
      RST     M653  ; 오3
      MPP
      OUT     T1997 K5
1499  LDP     T1997
      MOV     K8 D102
      ZP.PSTRT1 U7 D100 M100
1512  LD      M100
      ANI     M101
      OR      M436  ; 흡-
      AND     T1997
      OUT     M436  ; 흡-
1517  LD      X0A  ; 흡-
      OR      M437
      AND     M436  ; 흡-
      OUT     M437
1521  LDP     M437
      MOV     K9 D102
      ZP.PSTRT1 U7 D100 M100
1534  LD      M100
      ANI     M101
      OR      M438  ; 흡착OFFM2+
      AND     M437
      OUT     M438  ; 흡착OFFM2+
      OUT     T438 K5
      OUT     T439 K10
1547  LDP     T438
      MOV     K5 D102
      ZP.PSTRT1 U7 D100 M100
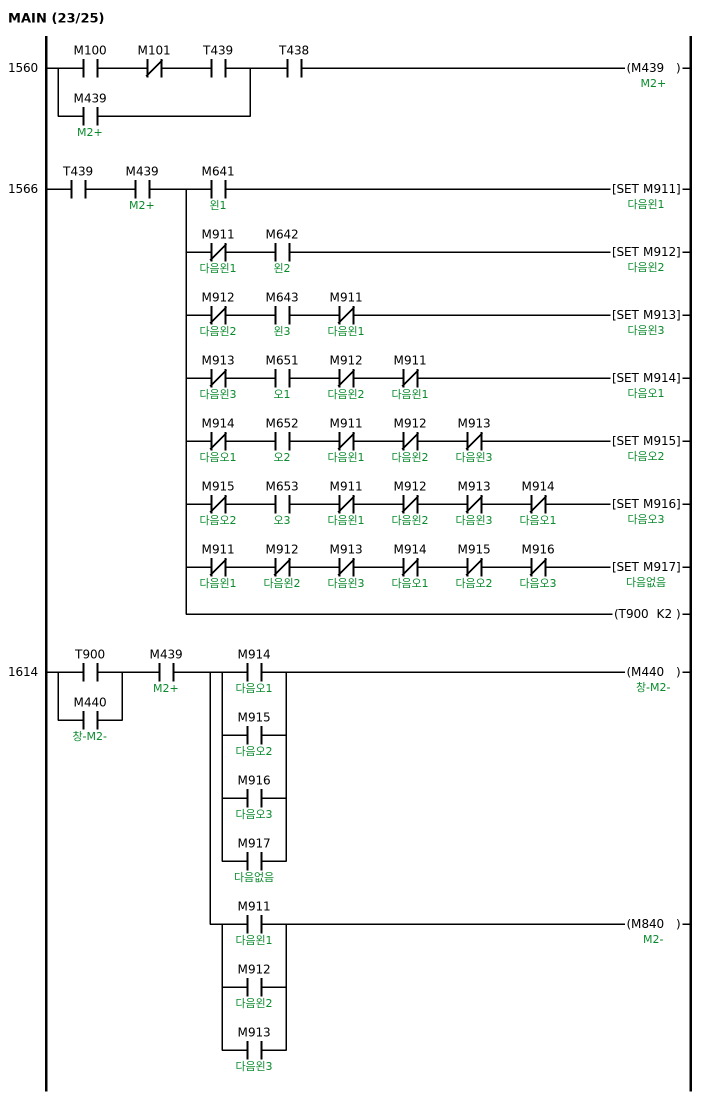
1560  LD      M100
      ANI     M101
      AND     T439
      OR      M439  ; M2+
      AND     T438
      OUT     M439  ; M2+
1566  LD      T439
      AND     M439  ; M2+
      MPS
      AND     M641  ; 왼1
      SET     M911  ; 다음왼1
      MRD
      ANI     M911  ; 다음왼1
      AND     M642  ; 왼2
      SET     M912  ; 다음왼2
      MRD
      ANI     M912  ; 다음왼2
      AND     M643  ; 왼3
      ANI     M911  ; 다음왼1
      SET     M913  ; 다음왼3
      MRD
      ANI     M913  ; 다음왼3
      AND     M651  ; 오1
      ANI     M912  ; 다음왼2
      ANI     M911  ; 다음왼1
      SET     M914  ; 다음오1
      MRD
      ANI     M914  ; 다음오1
      AND     M652  ; 오2
      ANI     M911  ; 다음왼1
      ANI     M912  ; 다음왼2
      ANI     M913  ; 다음왼3
      SET     M915  ; 다음오2
      MRD
      ANI     M915  ; 다음오2
      AND     M653  ; 오3
      ANI     M911  ; 다음왼1
      ANI     M912  ; 다음왼2
      ANI     M913  ; 다음왼3
      ANI     M914  ; 다음오1
      SET     M916  ; 다음오3
      MRD
      ANI     M911  ; 다음왼1
      ANI     M912  ; 다음왼2
      ANI     M913  ; 다음왼3
      ANI     M914  ; 다음오1
      ANI     M915  ; 다음오2
      ANI     M916  ; 다음오3
      SET     M917  ; 다음없음
      MPP
      OUT     T900 K2
1614  LD      T900
      OR      M440  ; 창-M2-
      AND     M439  ; M2+
      MPS
      LD      M914  ; 다음오1
      OR      M915  ; 다음오2
      OR      M916  ; 다음오3
      OR      M917  ; 다음없음
      ANB
      OUT     M440  ; 창-M2-
      MPP
      LD      M911  ; 다음왼1
      OR      M912  ; 다음왼2
      OR      M913  ; 다음왼3
      ANB
      OUT     M840  ; M2-
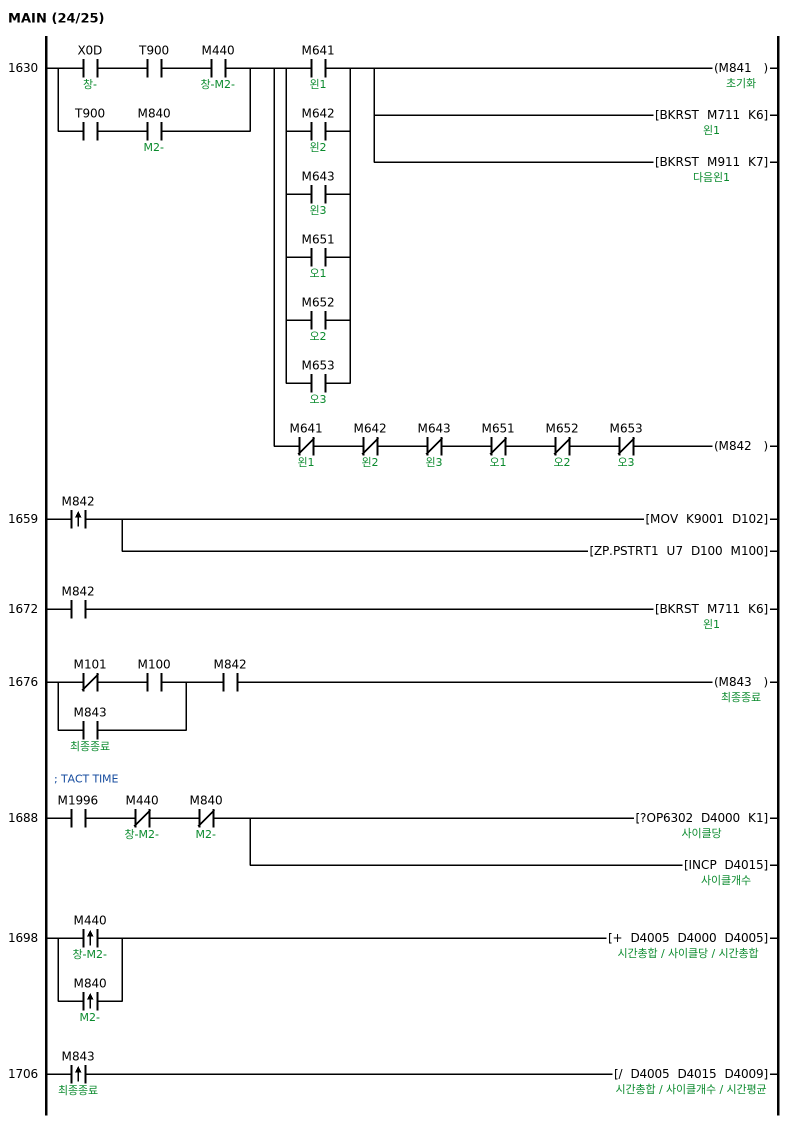
1630  LD      X0D  ; 창-
      AND     T900
      AND     M440  ; 창-M2-
      LD      T900
      AND     M840  ; M2-
      ORB
      MPS
      LD      M641  ; 왼1
      OR      M642  ; 왼2
      OR      M643  ; 왼3
      OR      M651  ; 오1
      OR      M652  ; 오2
      OR      M653  ; 오3
      ANB
      OUT     M841  ; 초기화
      BKRST   M711 K6
      BKRST   M911 K7
      MPP
      ANI     M641  ; 왼1
      ANI     M642  ; 왼2
      ANI     M643  ; 왼3
      ANI     M651  ; 오1
      ANI     M652  ; 오2
      ANI     M653  ; 오3
      OUT     M842
1659  LDP     M842
      MOV     K9001 D102
      ZP.PSTRT1 U7 D100 M100
1672  LD      M842
      BKRST   M711 K6
1676  LDI     M101
      AND     M100
      OR      M843  ; 최종종료
      AND     M842
      OUT     M843  ; 최종종료
; TACT TIME
1688  LD      M1996
      ANI     M440  ; 창-M2-
      ANI     M840  ; M2-
      ?OP6302 D4000 K1
      INCP    D4015
1698  LDP     M440  ; 창-M2-
      ORP     M840  ; M2-
      +       D4005 D4000 D4005
1706  LDP     M843  ; 최종종료
      /       D4005 D4015 D4009
